ABB RobotStudio station: Lab1_Decoracion.rsstn

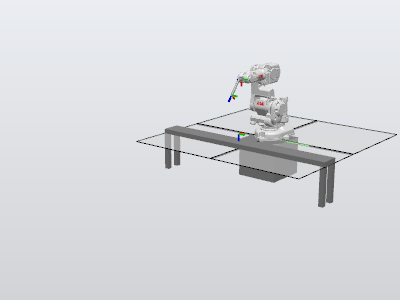
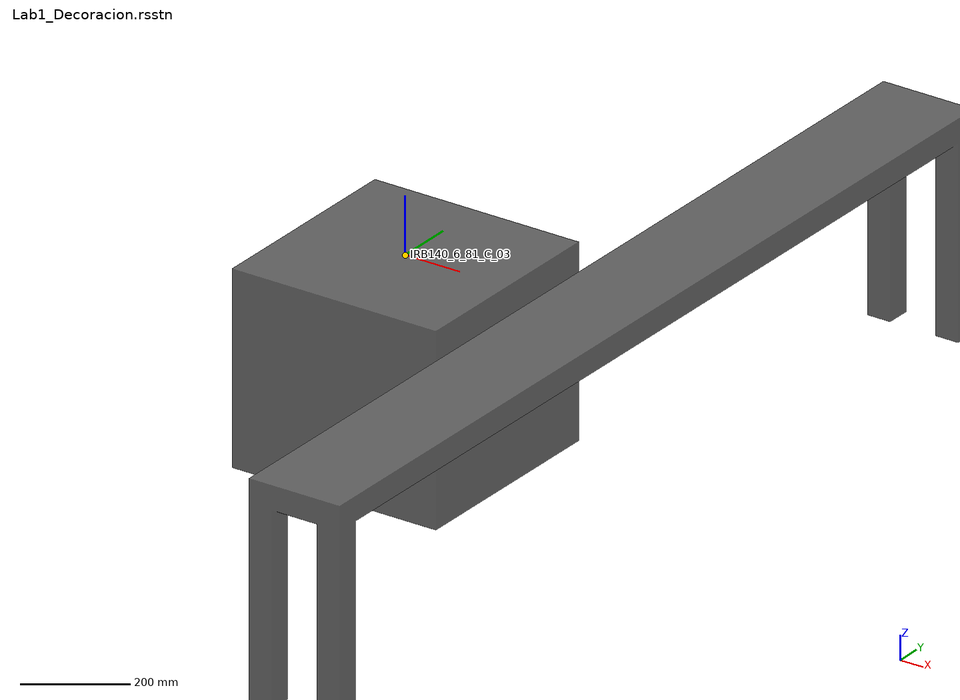
[picture v1: parts stored in the station drawn from their meshes, with robot base, taught points and paths (robot models come from the ABB library and are not in the file)]
Station Lab1_Decoracion (saved by RobotStudio 25.5.11605.0)
Controller Controlador_Lab1
  mechanical unit ROB_1: IRB140_6_81_C_03, 6 joints, base frame (0, 0, 0) mm
Layout (positions relative to the parent item):
  - IRB140_6_81_C_03 [mechanism, from %ABB.RobotStudio.Models.IRB140%\IRB140_6_81_C_G_03.rslib] at (0, 0, 0) mm; joint values [0, 0, 0, 0, 0, 0] (rad or m)
  - Pedestal [part] at (0, 0, -400) mm, size 450 x 450 x 400 mm
  - Banda_T [part] at (0, 0, -400) mm, size 200 x 2000 x 450 mm
  - Torta_1 [part] at (0, 0, -400) mm, size 240 x 240 x 115 mm
  - tool_Marcador [mechanism] at (515, 0, 712) mm, rotated rx 0 ry 90 rz 0 deg
      TCP tool_Marcador at (0, -139.3, 162.5) mm, rotated rx 0 ry 50 rz -90 deg
      links: ToolConMarcador_4
Attachment: tool_Marcador is attached to IRB140_6_81_C_03 / Link6
Targets, tools, work objects and paths stored in the station, written as RAPID:
! task T_ROB1
MODULE Mod_Decoracion
  PERS tooldata Tooldata_1:=[TRUE,[[139.3,0,162.5],[0.906307787,0,0.422618262,0]],[1,[52,0,82],[1,0,0,0],0,0,0]];
  PERS tooldata tool_Marcador:=[TRUE,[[139.3,0,162.5],[0.906307787,0,0.422618262,0]],[0.1,[52,0,82],[1,0,0,0],0,0,0]];
  TASK PERS wobjdata wobj_Torta:=[FALSE,TRUE,"",[[575,20,165],[0,0,1,0]],[[0,0,0],[1,0,0,0]]];
  PROC Prueba_Decoracion()
  ENDPROC
ENDMODULE

